TYPE ET_LeisterExtruder :
(
	ET_LeisterExtruder_eWaitExecute := 0,
	ET_LeisterExtruder_eStartExtruder,
	ET_LeisterExtruder_eStopExtruder,
	ET_LeisterExtruder_eWfHeaterReady,
	ET_LeisterExtruder_eDone := 197,
	ET_LeisterExtruder_eError := 198,
	ET_LeisterExtruder_eNoExecute := 199
);
END_TYPE

(* stored: Version 1.1.0.1, ProductVersion 3.1.4024.15
   DUT ET_LeisterExtruder: Id {da1ec206-4332-4aa4-94c2-3c78d2f17ce2} *)
